Fanuc KAREL source: KA00073.KL

PROGRAM KA00073
%NOLOCKGROUP
VAR
  SRC: XYZWPREXT
  DST: INTEGER
BEGIN
  SRC.X = 1.0
  DST = SRC
END KA00073
